Fanuc KAREL source: KT00551.KL

PROGRAM KT00551
%NOLOCKGROUP
VAR
  P1: JOINTPOS
  P2: JOINTPOS
  OUT: XYZWPREXT
BEGIN
  OUT = P1 : P2
END KT00551
